PROGRAM main
  VAR
    S1 AT %IX0.0  : BOOL; (* marcha / lote nuevo, NA *)
    S0 AT %IX0.1  : BOOL; (* parada, NC: TRUE sin pulsar *)
    B1 AT %IX0.2  : BOOL; (* sensor de piezas *)
    KM1 AT %QX0.0 : BOOL; (* motor de la cinta *)
    H1 AT %QX0.1  : BOOL; (* lote completo *)
    F_PIEZA       : R_TRIG;
    PIEZAS        : INT; (* piezas del lote *)
    COMPLETO      : BOOL; (* lote completo *)
    F_LOTE        : R_TRIG;
    LOTES         : INT; (* lotes completos en el turno *)
    TURNO         : BOOL; (* turno completo *)
  END_VAR
  VAR  (* added by the conversion: wires and edge detectors of the diagram *)
    R_TRIG1 : R_TRIG;
    R_TRIG2 : R_TRIG;
  END_VAR

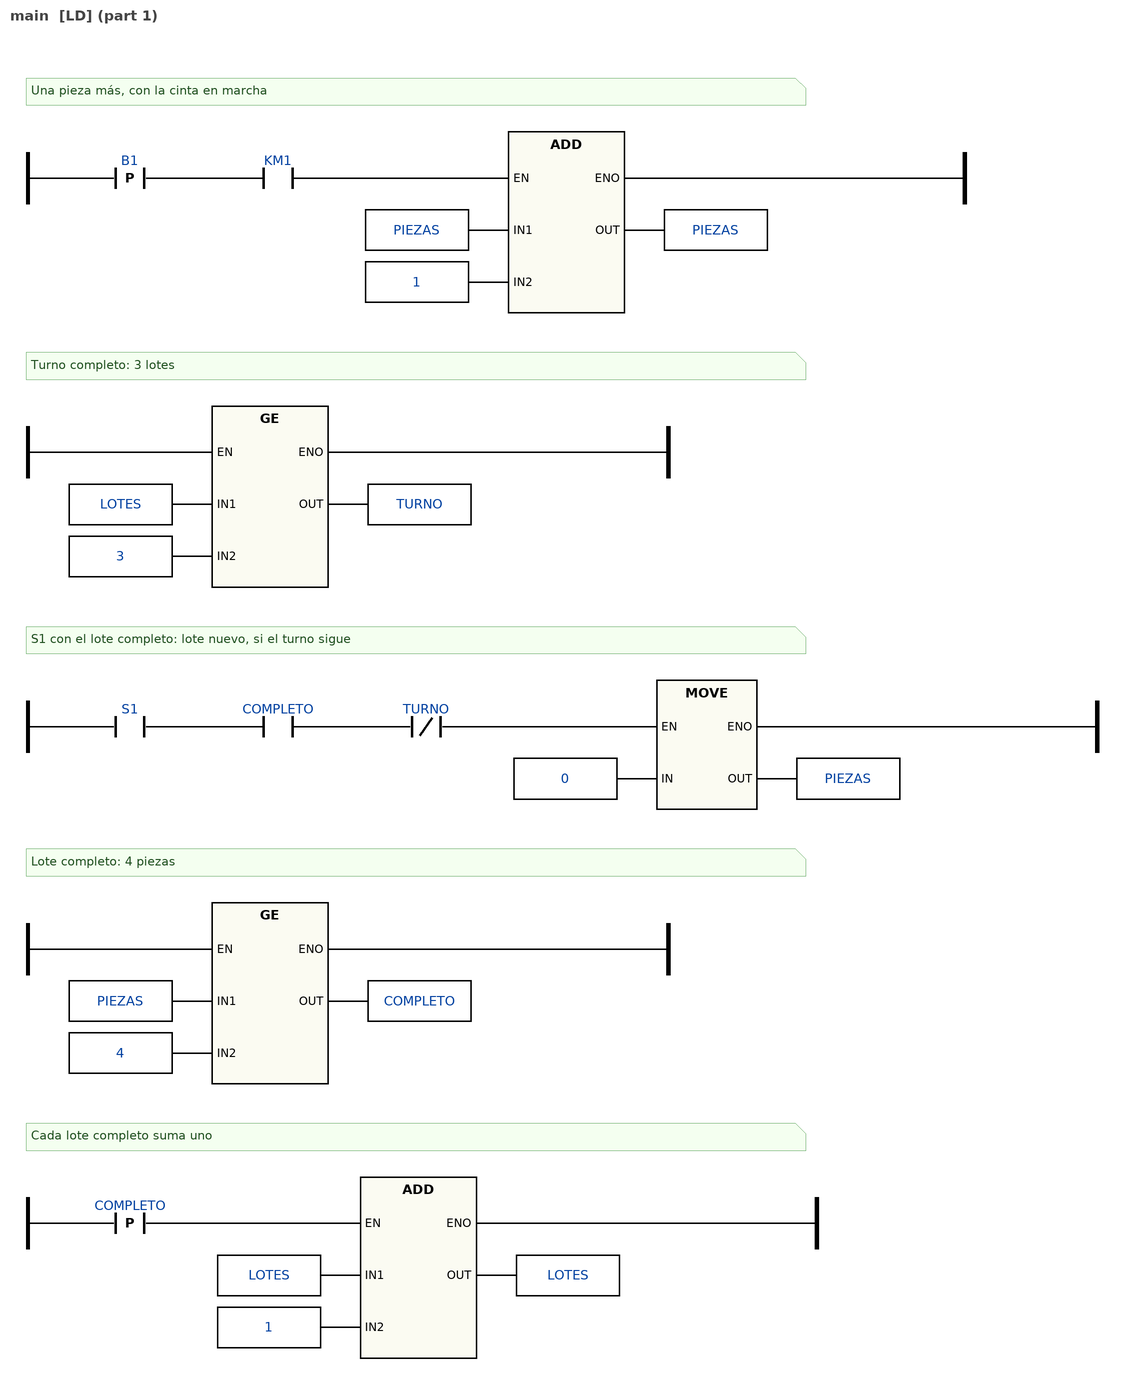
(* LD diagram, written out as Structured Text *)
(* Una pieza más, con la cinta en marcha *)
R_TRIG1(CLK := B1);
IF R_TRIG1.Q AND KM1 THEN PIEZAS := PIEZAS + 1; END_IF;
(* Turno completo: 3 lotes *)
TURNO := LOTES >= 3;
(* S1 con el lote completo: lote nuevo, si el turno sigue *)
IF S1 AND COMPLETO AND NOT TURNO THEN PIEZAS := 0; END_IF;
(* Lote completo: 4 piezas *)
COMPLETO := PIEZAS >= 4;
(* Cada lote completo suma uno *)
R_TRIG2(CLK := COMPLETO);
IF R_TRIG2.Q THEN LOTES := LOTES + 1; END_IF;
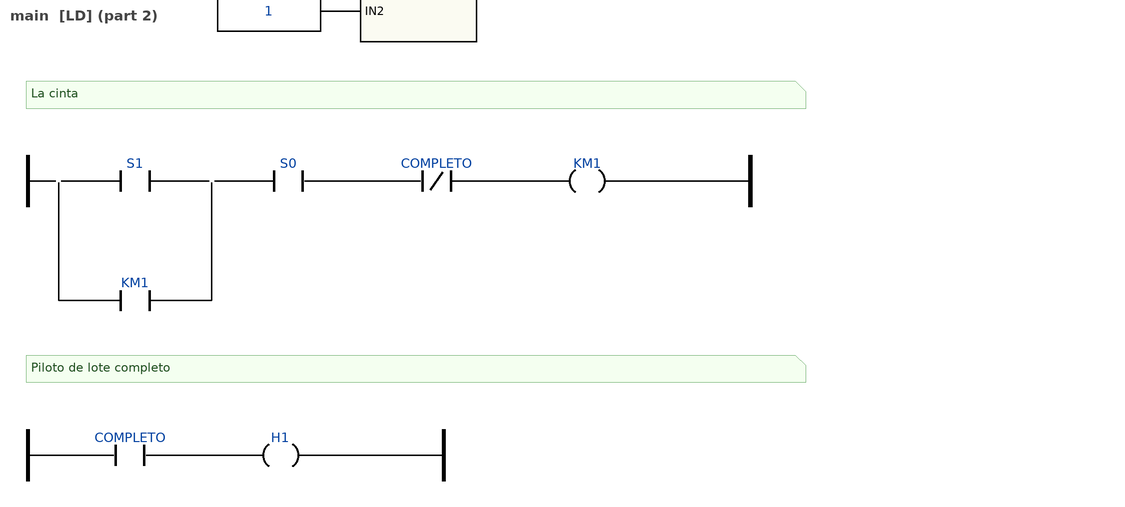
(* La cinta *)
KM1 := (S1 OR KM1) AND S0 AND NOT COMPLETO;
(* Piloto de lote completo *)
H1 := COMPLETO;
END_PROGRAM
